// TIA Portal V20 export
// export: Created 2026-10-20T12:51:09.2669842Z, ExportSetting WithDefaults, DisplayName Totally Integrated Automation Portal, DisplayVersion V20 Update 6, DisplayName TIA Portal Openness, DisplayVersion V20 Update 6, DisplayName TIA Portal Version Control Interface, DisplayVersion V20 Update 6, DisplayName SINAMICS Startdrive Advanced, DisplayVersion V20 SP1, DisplayName SINAMICS Startdrive G130, G150, S120, S150, SINAMICS MV, G220, S200, S210, DisplayVersion V20 SP1, DisplayName SINAMICS Startdrive G110M, G120, G120C, G120D, G120P, G115D, DisplayVersion V20 SP1, DisplayName STEP 7 Professional, DisplayVersion V20 Update 6, DisplayName STEP 7 Safety, DisplayVersion V20 Update 2, DisplayName WinCC Basic/Comfort/Advanced, DisplayVersion V20 Update 6, DisplayName WinCC Unified, DisplayVersion V20 Update 6
FUNCTION_BLOCK "Remote_Panel"   // FB17, F_LAD
{ S7_Optimized_Access := 'TRUE' }
VERSION : 0.1
// stored: AutoNumber true, IsIECCheckEnabled false, UDAEnableTagReadback false
   VAR_INPUT
      ID : Int;
      Overtravel_Lower_limit : Bool;
      Overtravel_Upper_limit : Bool;
      Estop : Bool;
      Reset : Bool;
      Chain_Slack_1 : Bool;
      Chain_Slack_2 : Bool;
      Chain_Slack_3 : Bool;
      Chain_Slack_4 : Bool;
      "Light Guards CX101" : Bool;
      "Light Guards CX201" : Bool;
      Gate_1 : Bool;
      Gate_2 : Bool;
      EStop_Lock_1 : Bool;
      EStop_Lock_2 : Bool;
      Lock_Secured_1 : Bool;
      Lock_Secured_2 : Bool;
      "EStop Level 1" : Bool;
      "EStop Level 2" : Bool;
      "EStop Level 3" : Bool;
      "EStop Level 4" : Bool;
      "EStop Level 5" : Bool;
      "EStop Level 6" : Bool;
      "EStop Level 7" : Bool;
      "EStop Level 8" : Bool;
      Bypass : "F_Bypass_RemotePanel";
      Material_Selection_1 : Bool;
      MR_1 : Bool;
      Material_Selection_2 : Bool;
      MR_2 : Bool;
      Overhang_Left : Bool;
      Overhang_Right : Bool;
   END_VAR
   VAR_OUTPUT
      Safety_OK : Bool;
      Bypass_Warning : Bool;
      "STO VTD - CH1" : Bool;
      "STO VTD - CH2" : Bool;
      "STO CONVEYOR VTD - CH1" : Bool;
      "STO CONVEYOR VTD - CH2" : Bool;
      "STO CNV VFD (Level 1,2,3 - Side1) - CH1" : Bool;
      "STO CNV VFD (Level 1,2,3 - Side1) - CH2" : Bool;
      "STO CNV VFD (Level 1,2,3 - Side2) - CH1" : Bool;
      "STO CNV VFD (Level 1,2,3 - Side2) - CH2" : Bool;
      "STO CNV VFD (Level 4,5,6 - Side1) - CH1" : Bool;
      "STO CNV VFD (Level 4,5,6 - Side1) - CH2" : Bool;
      "STO CNV VFD (Level 4,5,6 - Side2) - CH1" : Bool;
      "STO CNV VFD (Level 4,5,6 - Side2) - CH2" : Bool;
      "STO CNV VFD (Level 7,8 - Side1) - CH1" : Bool;
      "STO CNV VFD (Level 7,8 - Side1) - CH2" : Bool;
      "STO CNV VFD (Level 7,8 - Side2) - CH1" : Bool;
      "STO CNV VFD (Level 7,8 - Side2) - CH2" : Bool;
      "Power Enable Safety Stopper Conveyors (Level 1,2,3 - Side1) - CH1" : Bool;
      "Power Enable Safety Stopper Conveyors (Level 1,2,3 - Side1) - CH2" : Bool;
      "Power Enable Safety Stopper Conveyors (Level 1,2,3 - Side2) - CH1" : Bool;
      "Power Enable Safety Stopper Conveyors (Level 1,2,3 - Side2) - CH2" : Bool;
      "Power Enable Safety Stopper Conveyors (Level 4,5,6 - Side1) - CH1" : Bool;
      "Power Enable Safety Stopper Conveyors (Level 4,5,6 - Side1) - CH2" : Bool;
      "Power Enable Safety Stopper Conveyors (Level 4,5,6 - Side2) - CH1" : Bool;
      "Power Enable Safety Stopper Conveyors (Level 4,5,6 - Side2) - CH2" : Bool;
      "Power Enable Safety Stopper Conveyors (Level 7,8 - Side1) - CH1" : Bool;
      "Power Enable Safety Stopper Conveyors (Level 7,8 - Side1) - CH2" : Bool;
      "Power Enable Safety Stopper Conveyors (Level 7,8 - Side2) - CH1" : Bool;
      "Power Enable Safety Stopper Conveyors (Level 7,8 - Side2) - CH2" : Bool;
      "VTU Hoist Brake Sfty Enable - CH1" : Bool;
      "VTU Hoist Brake Sfty Enable - CH2" : Bool;
      ACK { ExternalAccessible := 'False'; ExternalVisible := 'False'; ExternalWritable := 'False'} : Bool;
      L1_OK : Bool;
      L2_OK : Bool;
      L3_OK : Bool;
      L4_OK : Bool;
      L5_OK : Bool;
      L6_OK : Bool;
      L7_OK : Bool;
      L8_OK : Bool;
      EStop_Lock_1_OK : Bool;
      EStop_Lock_2_OK : Bool;
      Lock_Secured_1_OK : Bool;
      Lock_Secured_2_OK : Bool;
      Safety_Ok_Conf : Bool;
   END_VAR
   VAR
      Overtravel_Lower_Limit_DB : ESTOP1;
      Overtravel_Upper_Limit_DB : ESTOP1;
      Estop_Cabinet_DB : ESTOP1;
      Chain_Slack_1_DB : ESTOP1;
      Chain_Slack_2_DB : ESTOP1;
      Chain_Slack_3_DB : ESTOP1;
      Chain_Slack_4_DB : ESTOP1;
      Light_Guards_CX101 : ESTOP1;
      Light_Guards_CX201 : ESTOP1;
      Gate_1_DB : ESTOP1;
      Gate_2_DB : ESTOP1;
      EStop_Lock_1_DB : ESTOP1;
      EStop_Lock_2_DB : ESTOP1;
      Lock_Secured_1_DB : ESTOP1;
      Lock_Secured_2_DB : ESTOP1;
      "EStop Level 1_DB" : ESTOP1;
      "EStop Level 2_DB" : ESTOP1;
      "EStop Level 3_DB" : ESTOP1;
      "EStop Level 4_DB" : ESTOP1;
      "EStop Level 5_DB" : ESTOP1;
      "EStop Level 6_DB" : ESTOP1;
      "EStop Level 7_DB" : ESTOP1;
      "EStop Level 8_DB" : ESTOP1;
      Mute_LG_1_DB : "SICK Safe Entry Exit HW PLC V02";
      Distance_Materia_To_LG : DInt;
      Mute_LG_2_DB : "SICK Safe Entry Exit HW PLC V02";
      F_T_Delay_Sae_OK : TOF;
      F_T_Delay_CL_4 : TOF;
      F_T_Delay_CL_3 : TOF;
      F_T_Delay_CL_2 : TOF;
      F_T_Delay_CL_1 : TOF;
      Chain_Slack_1_Filtered { ExternalAccessible := 'False'; ExternalVisible := 'False'; ExternalWritable := 'False'} : Bool;
      Chain_Slack_2_Filtered { ExternalAccessible := 'False'; ExternalVisible := 'False'; ExternalWritable := 'False'} : Bool;
      Chain_Slack_3_Filtered { ExternalAccessible := 'False'; ExternalVisible := 'False'; ExternalWritable := 'False'} : Bool;
      Chain_Slack_4_Filtered { ExternalAccessible := 'False'; ExternalVisible := 'False'; ExternalWritable := 'False'} : Bool;
      Light_Guard_Tuned : Bool;
      Light_Guard_Tuned_Euro : Bool;
      Light_Guard_Tuned_UK : Bool;
      Light_Guard_Tuned_UK_Infeed : Bool;
      Light_Guard_Tuned_Euro_Infeed : Bool;
      Light_Guard_Tuned_Infeed : Bool;
      F_Timer_Infeed_UK : TP;
      F_Timer_Infeed_E : TP;
      F_Timer_Outfeed_UK : TP;
      F_Timer_Outfeed_E : TP;
      Overhang_Left_DB : ESTOP1;
      Overhang_Right_DB : ESTOP1;
   END_VAR
   VAR_TEMP
      EStop_Levels_OK : Bool;
   END_VAR
   VAR_TEMP   // added for the SCL form of the ladder/FBD networks
      _w1 : Bool;
   END_VAR
BEGIN

REGION Network 1: RESET CABINET
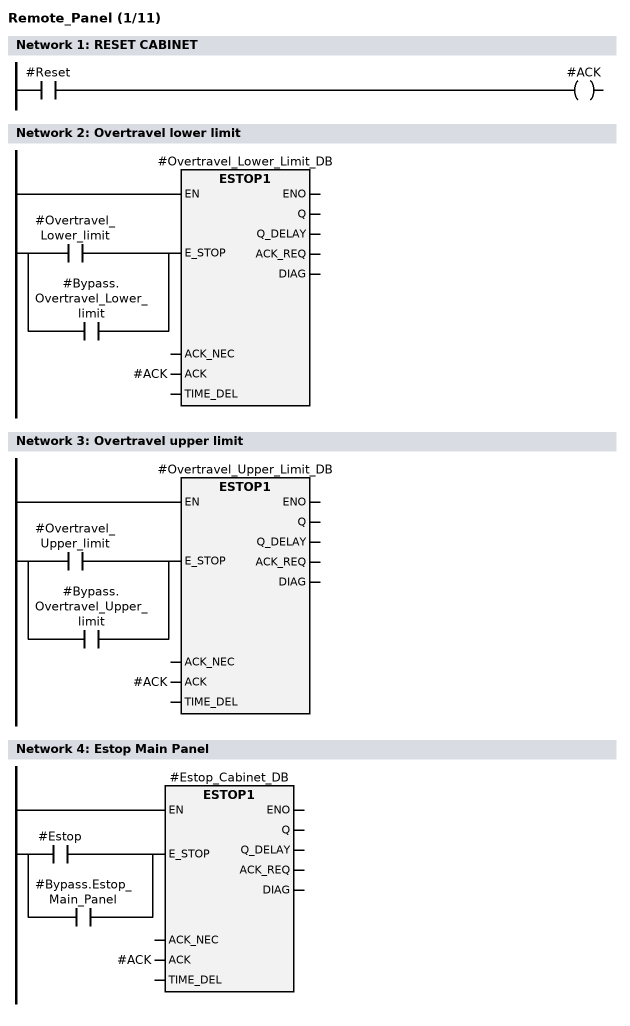
   RUNG wire#powerrail
      Contact( #Reset )
      Coil( #ACK )
   END_RUNG
   // the same network as SCL:
   #ACK := #Reset;
END_REGION

REGION Network 2: Overtravel lower limit
   RUNG wire#powerrail
      #Overtravel_Lower_Limit_DB.ESTOP1(E_STOP := wire#w1, ACK_NEC :=, ACK := #ACK, TIME_DEL :=, Q =>, Q_DELAY =>, ACK_REQ =>, DIAG =>)
   END_RUNG
   RUNG wire#powerrail
      Contact( #Overtravel_Lower_limit )
   END_RUNG wire#w1
   RUNG wire#powerrail
      Contact( #Bypass.Overtravel_Lower_limit )
   END_RUNG wire#w1
   // the same network as SCL:
   #Overtravel_Lower_Limit_DB(E_STOP := #Overtravel_Lower_limit OR #Bypass.Overtravel_Lower_limit, ACK := #ACK);   // ESTOP1
END_REGION

REGION Network 3: Overtravel upper limit
   RUNG wire#powerrail
      #Overtravel_Upper_Limit_DB.ESTOP1(E_STOP := wire#w1, ACK_NEC :=, ACK := #ACK, TIME_DEL :=, Q =>, Q_DELAY =>, ACK_REQ =>, DIAG =>)
   END_RUNG
   RUNG wire#powerrail
      Contact( #Overtravel_Upper_limit )
   END_RUNG wire#w1
   RUNG wire#powerrail
      Contact( #Bypass.Overtravel_Upper_limit )
   END_RUNG wire#w1
   // the same network as SCL:
   #Overtravel_Upper_Limit_DB(E_STOP := #Overtravel_Upper_limit OR #Bypass.Overtravel_Upper_limit, ACK := #ACK);   // ESTOP1
END_REGION

REGION Network 4: Estop Main Panel
   RUNG wire#powerrail
      #Estop_Cabinet_DB.ESTOP1(E_STOP := wire#w1, ACK_NEC :=, ACK := #ACK, TIME_DEL :=, Q =>, Q_DELAY =>, ACK_REQ =>, DIAG =>)
   END_RUNG
   RUNG wire#powerrail
      Contact( #Estop )
   END_RUNG wire#w1
   RUNG wire#powerrail
      Contact( #Bypass.Estop_Main_Panel )
   END_RUNG wire#w1
   // the same network as SCL:
   #Estop_Cabinet_DB(E_STOP := #Estop OR #Bypass.Estop_Main_Panel, ACK := #ACK);   // ESTOP1
END_REGION

REGION Network 5: Chain slack 1
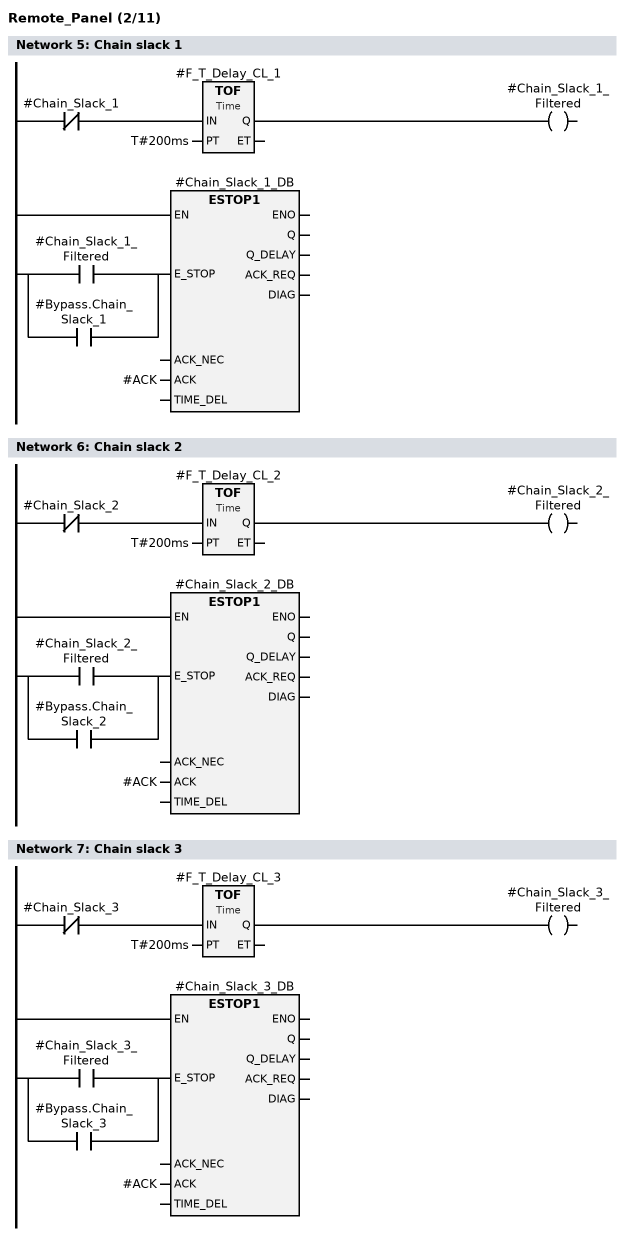
   RUNG wire#powerrail
      I_Contact( #Chain_Slack_1 )
      { S7_Templates := "[time_type := Time, codedbool_type := DInt]" } #F_T_Delay_CL_1.TOF(pt := T#200ms, et =>)
      Coil( #Chain_Slack_1_Filtered )
   END_RUNG
   RUNG wire#powerrail
      #Chain_Slack_1_DB.ESTOP1(E_STOP := wire#w1, ACK_NEC :=, ACK := #ACK, TIME_DEL :=, Q =>, Q_DELAY =>, ACK_REQ =>, DIAG =>)
   END_RUNG
   RUNG wire#powerrail
      Contact( #Chain_Slack_1_Filtered )
   END_RUNG wire#w1
   RUNG wire#powerrail
      Contact( #Bypass.Chain_Slack_1 )
   END_RUNG wire#w1
   // the same network as SCL:
   #F_T_Delay_CL_1.TOF(IN := NOT #Chain_Slack_1, PT := T#200ms);
   #Chain_Slack_1_Filtered := #F_T_Delay_CL_1.Q;
   #Chain_Slack_1_DB(E_STOP := #Chain_Slack_1_Filtered OR #Bypass.Chain_Slack_1, ACK := #ACK);   // ESTOP1
END_REGION

REGION Network 6: Chain slack 2
   RUNG wire#powerrail
      I_Contact( #Chain_Slack_2 )
      { S7_Templates := "[time_type := Time, codedbool_type := DInt]" } #F_T_Delay_CL_2.TOF(pt := T#200ms, et =>)
      Coil( #Chain_Slack_2_Filtered )
   END_RUNG
   RUNG wire#powerrail
      #Chain_Slack_2_DB.ESTOP1(E_STOP := wire#w1, ACK_NEC :=, ACK := #ACK, TIME_DEL :=, Q =>, Q_DELAY =>, ACK_REQ =>, DIAG =>)
   END_RUNG
   RUNG wire#powerrail
      Contact( #Chain_Slack_2_Filtered )
   END_RUNG wire#w1
   RUNG wire#powerrail
      Contact( #Bypass.Chain_Slack_2 )
   END_RUNG wire#w1
   // the same network as SCL:
   #F_T_Delay_CL_2.TOF(IN := NOT #Chain_Slack_2, PT := T#200ms);
   #Chain_Slack_2_Filtered := #F_T_Delay_CL_2.Q;
   #Chain_Slack_2_DB(E_STOP := #Chain_Slack_2_Filtered OR #Bypass.Chain_Slack_2, ACK := #ACK);   // ESTOP1
END_REGION

REGION Network 7: Chain slack 3
   RUNG wire#powerrail
      I_Contact( #Chain_Slack_3 )
      { S7_Templates := "[time_type := Time, codedbool_type := DInt]" } #F_T_Delay_CL_3.TOF(pt := T#200ms, et =>)
      Coil( #Chain_Slack_3_Filtered )
   END_RUNG
   RUNG wire#powerrail
      #Chain_Slack_3_DB.ESTOP1(E_STOP := wire#w1, ACK_NEC :=, ACK := #ACK, TIME_DEL :=, Q =>, Q_DELAY =>, ACK_REQ =>, DIAG =>)
   END_RUNG
   RUNG wire#powerrail
      Contact( #Chain_Slack_3_Filtered )
   END_RUNG wire#w1
   RUNG wire#powerrail
      Contact( #Bypass.Chain_Slack_3 )
   END_RUNG wire#w1
   // the same network as SCL:
   #F_T_Delay_CL_3.TOF(IN := NOT #Chain_Slack_3, PT := T#200ms);
   #Chain_Slack_3_Filtered := #F_T_Delay_CL_3.Q;
   #Chain_Slack_3_DB(E_STOP := #Chain_Slack_3_Filtered OR #Bypass.Chain_Slack_3, ACK := #ACK);   // ESTOP1
END_REGION

REGION Network 8: Chain slack 4
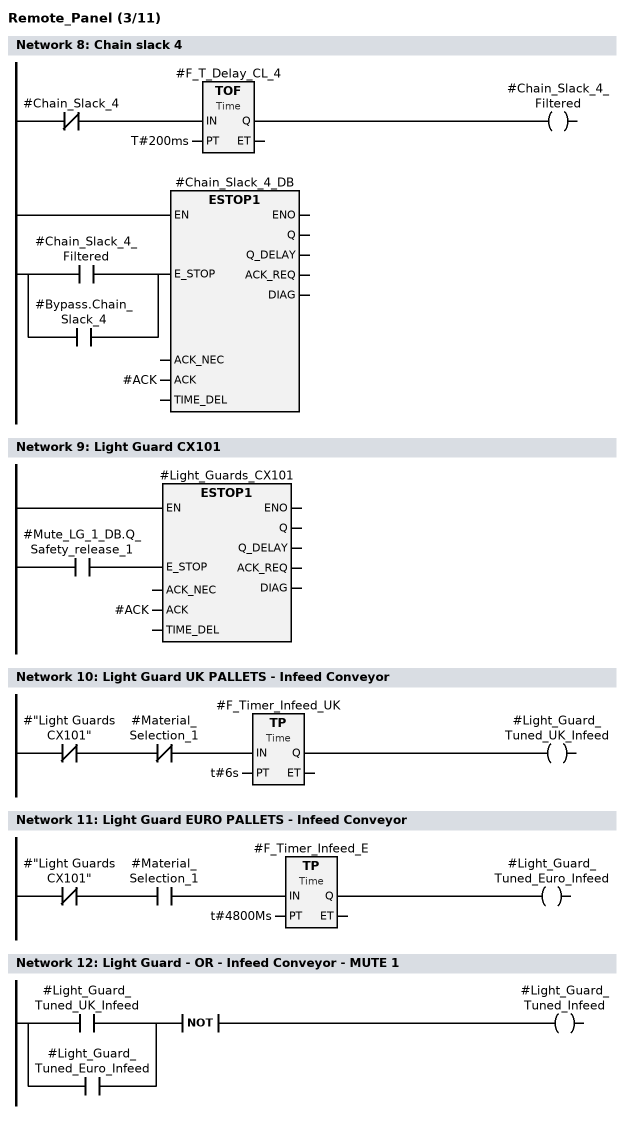
   RUNG wire#powerrail
      I_Contact( #Chain_Slack_4 )
      { S7_Templates := "[time_type := Time, codedbool_type := DInt]" } #F_T_Delay_CL_4.TOF(pt := T#200ms, et =>)
      Coil( #Chain_Slack_4_Filtered )
   END_RUNG
   RUNG wire#powerrail
      #Chain_Slack_4_DB.ESTOP1(E_STOP := wire#w1, ACK_NEC :=, ACK := #ACK, TIME_DEL :=, Q =>, Q_DELAY =>, ACK_REQ =>, DIAG =>)
   END_RUNG
   RUNG wire#powerrail
      Contact( #Chain_Slack_4_Filtered )
   END_RUNG wire#w1
   RUNG wire#powerrail
      Contact( #Bypass.Chain_Slack_4 )
   END_RUNG wire#w1
   // the same network as SCL:
   #F_T_Delay_CL_4.TOF(IN := NOT #Chain_Slack_4, PT := T#200ms);
   #Chain_Slack_4_Filtered := #F_T_Delay_CL_4.Q;
   #Chain_Slack_4_DB(E_STOP := #Chain_Slack_4_Filtered OR #Bypass.Chain_Slack_4, ACK := #ACK);   // ESTOP1
END_REGION

REGION Network 9: Light Guard CX101
   RUNG wire#powerrail
      #Light_Guards_CX101.ESTOP1(E_STOP := wire#w1, ACK_NEC :=, ACK := #ACK, TIME_DEL :=, Q =>, Q_DELAY =>, ACK_REQ =>, DIAG =>)
   END_RUNG
   RUNG wire#powerrail
      Contact( #Mute_LG_1_DB.Q_Safety_release_1 )
   END_RUNG wire#w1
   // the same network as SCL:
   #Light_Guards_CX101(E_STOP := #Mute_LG_1_DB.Q_Safety_release_1, ACK := #ACK);   // ESTOP1
END_REGION

REGION Network 10: Light Guard UK PALLETS - Infeed Conveyor
   RUNG wire#powerrail
      I_Contact( #"Light Guards CX101" )
      I_Contact( #Material_Selection_1 )
      { S7_Templates := "[time_type := Time, codedbool_type := DInt]" } #F_Timer_Infeed_UK.TP(pt := t#6s, et =>)
      Coil( #Light_Guard_Tuned_UK_Infeed )
   END_RUNG
   // the same network as SCL:
   #F_Timer_Infeed_UK.TP(IN := NOT #"Light Guards CX101" AND NOT #Material_Selection_1, PT := t#6s);
   #Light_Guard_Tuned_UK_Infeed := #F_Timer_Infeed_UK.Q;
END_REGION

REGION Network 11: Light Guard EURO PALLETS - Infeed Conveyor
   RUNG wire#powerrail
      I_Contact( #"Light Guards CX101" )
      Contact( #Material_Selection_1 )
      { S7_Templates := "[time_type := Time, codedbool_type := DInt]" } #F_Timer_Infeed_E.TP(pt := t#4800Ms, et =>)
      Coil( #Light_Guard_Tuned_Euro_Infeed )
   END_RUNG
   // the same network as SCL:
   #F_Timer_Infeed_E.TP(IN := NOT #"Light Guards CX101" AND #Material_Selection_1, PT := t#4800Ms);
   #Light_Guard_Tuned_Euro_Infeed := #F_Timer_Infeed_E.Q;
END_REGION

REGION Network 12: Light Guard - OR - Infeed Conveyor - MUTE 1
   RUNG wire#powerrail
      Contact( #Light_Guard_Tuned_UK_Infeed )
      wire#w1
      Not()
      Coil( #Light_Guard_Tuned_Infeed )
   END_RUNG
   RUNG wire#powerrail
      Contact( #Light_Guard_Tuned_Euro_Infeed )
   END_RUNG wire#w1
   // the same network as SCL:
   #Light_Guard_Tuned_Infeed := NOT (#Light_Guard_Tuned_UK_Infeed OR #Light_Guard_Tuned_Euro_Infeed);
END_REGION

REGION Network 13: MUTE 1
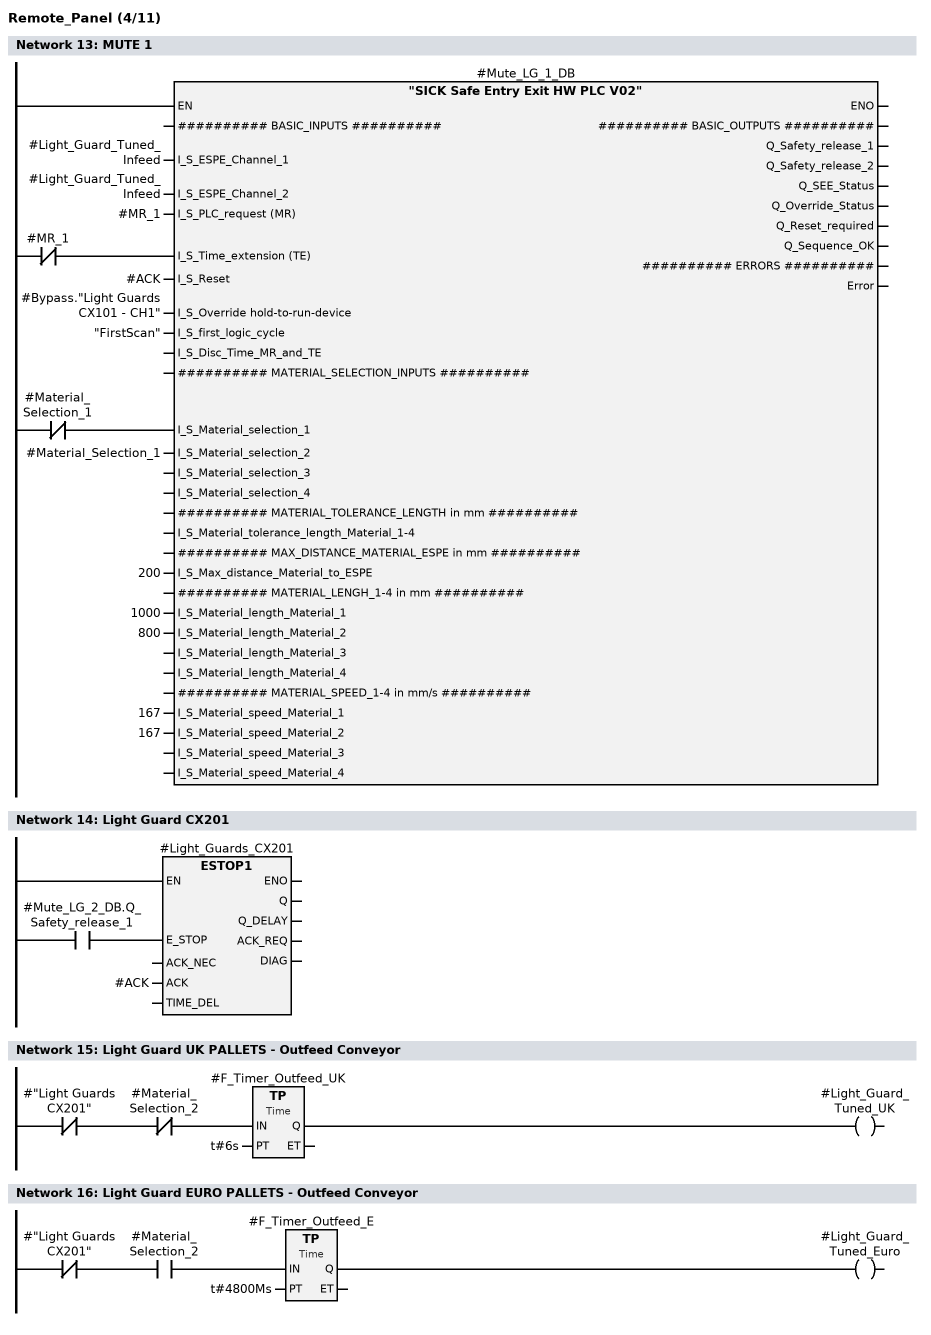
   RUNG wire#powerrail
      #Mute_LG_1_DB("I_S_Time_extension (TE)" := wire#w1, I_S_Material_selection_1 := wire#w2, "########## BASIC_INPUTS ##########" :=, I_S_ESPE_Channel_1 := #Light_Guard_Tuned_Infeed, I_S_ESPE_Channel_2 := #Light_Guard_Tuned_Infeed, "I_S_PLC_request (MR)" := #MR_1, I_S_Reset := #ACK, "I_S_Override hold-to-run-device" := #Bypass."Light Guards CX101 - CH1", I_S_first_logic_cycle := "FirstScan", I_S_Disc_Time_MR_and_TE :=, "########## MATERIAL_SELECTION_INPUTS ##########" :=, I_S_Material_selection_2 := #Material_Selection_1, I_S_Material_selection_3 :=, I_S_Material_selection_4 :=, "########## MATERIAL_TOLERANCE_LENGTH in mm ##########" :=, "I_S_Material_tolerance_length_Material_1-4" :=, "########## MAX_DISTANCE_MATERIAL_ESPE in mm ##########" :=, I_S_Max_distance_Material_to_ESPE := 200, "########## MATERIAL_LENGH_1-4 in mm ##########" :=, I_S_Material_length_Material_1 := 1000, I_S_Material_length_Material_2 := 800, I_S_Material_length_Material_3 :=, I_S_Material_length_Material_4 :=, "########## MATERIAL_SPEED_1-4 in mm/s ##########" :=, I_S_Material_speed_Material_1 := 167, I_S_Material_speed_Material_2 := 167, I_S_Material_speed_Material_3 :=, I_S_Material_speed_Material_4 :=, "########## BASIC_OUTPUTS ##########" =>, Q_Safety_release_1 =>, Q_Safety_release_2 =>, Q_SEE_Status =>, Q_Override_Status =>, Q_Reset_required =>, Q_Sequence_OK =>, "########## ERRORS ##########" =>, Error =>)
   END_RUNG
   RUNG wire#powerrail
      I_Contact( #MR_1 )
   END_RUNG wire#w1
   RUNG wire#powerrail
      I_Contact( #Material_Selection_1 )
   END_RUNG wire#w2
   // the same network as SCL:
   #Mute_LG_1_DB(I_S_ESPE_Channel_1 := #Light_Guard_Tuned_Infeed,   // "SICK Safe Entry Exit HW PLC V02"
                 I_S_ESPE_Channel_2 := #Light_Guard_Tuned_Infeed,
                 "I_S_PLC_request (MR)" := #MR_1,
                 "I_S_Time_extension (TE)" := NOT #MR_1,
                 I_S_Reset := #ACK,
                 "I_S_Override hold-to-run-device" := #Bypass."Light Guards CX101 - CH1",
                 I_S_first_logic_cycle := "FirstScan",
                 I_S_Material_selection_1 := NOT #Material_Selection_1,
                 I_S_Material_selection_2 := #Material_Selection_1,
                 I_S_Max_distance_Material_to_ESPE := 200,
                 I_S_Material_length_Material_1 := 1000,
                 I_S_Material_length_Material_2 := 800,
                 I_S_Material_speed_Material_1 := 167,
                 I_S_Material_speed_Material_2 := 167);
END_REGION

REGION Network 14: Light Guard CX201
   RUNG wire#powerrail
      #Light_Guards_CX201.ESTOP1(E_STOP := wire#w1, ACK_NEC :=, ACK := #ACK, TIME_DEL :=, Q =>, Q_DELAY =>, ACK_REQ =>, DIAG =>)
   END_RUNG
   RUNG wire#powerrail
      Contact( #Mute_LG_2_DB.Q_Safety_release_1 )
   END_RUNG wire#w1
   // the same network as SCL:
   #Light_Guards_CX201(E_STOP := #Mute_LG_2_DB.Q_Safety_release_1, ACK := #ACK);   // ESTOP1
END_REGION

REGION Network 15: Light Guard UK PALLETS - Outfeed Conveyor
   RUNG wire#powerrail
      I_Contact( #"Light Guards CX201" )
      I_Contact( #Material_Selection_2 )
      { S7_Templates := "[time_type := Time, codedbool_type := DInt]" } #F_Timer_Outfeed_UK.TP(pt := t#6s, et =>)
      Coil( #Light_Guard_Tuned_UK )
   END_RUNG
   // the same network as SCL:
   #F_Timer_Outfeed_UK.TP(IN := NOT #"Light Guards CX201" AND NOT #Material_Selection_2, PT := t#6s);
   #Light_Guard_Tuned_UK := #F_Timer_Outfeed_UK.Q;
END_REGION

REGION Network 16: Light Guard EURO PALLETS - Outfeed Conveyor
   RUNG wire#powerrail
      I_Contact( #"Light Guards CX201" )
      Contact( #Material_Selection_2 )
      { S7_Templates := "[time_type := Time, codedbool_type := DInt]" } #F_Timer_Outfeed_E.TP(pt := t#4800Ms, et =>)
      Coil( #Light_Guard_Tuned_Euro )
   END_RUNG
   // the same network as SCL:
   #F_Timer_Outfeed_E.TP(IN := NOT #"Light Guards CX201" AND #Material_Selection_2, PT := t#4800Ms);
   #Light_Guard_Tuned_Euro := #F_Timer_Outfeed_E.Q;
END_REGION

REGION Network 17: Light Guard - OR - Infeed Conveyor - MUTE 2
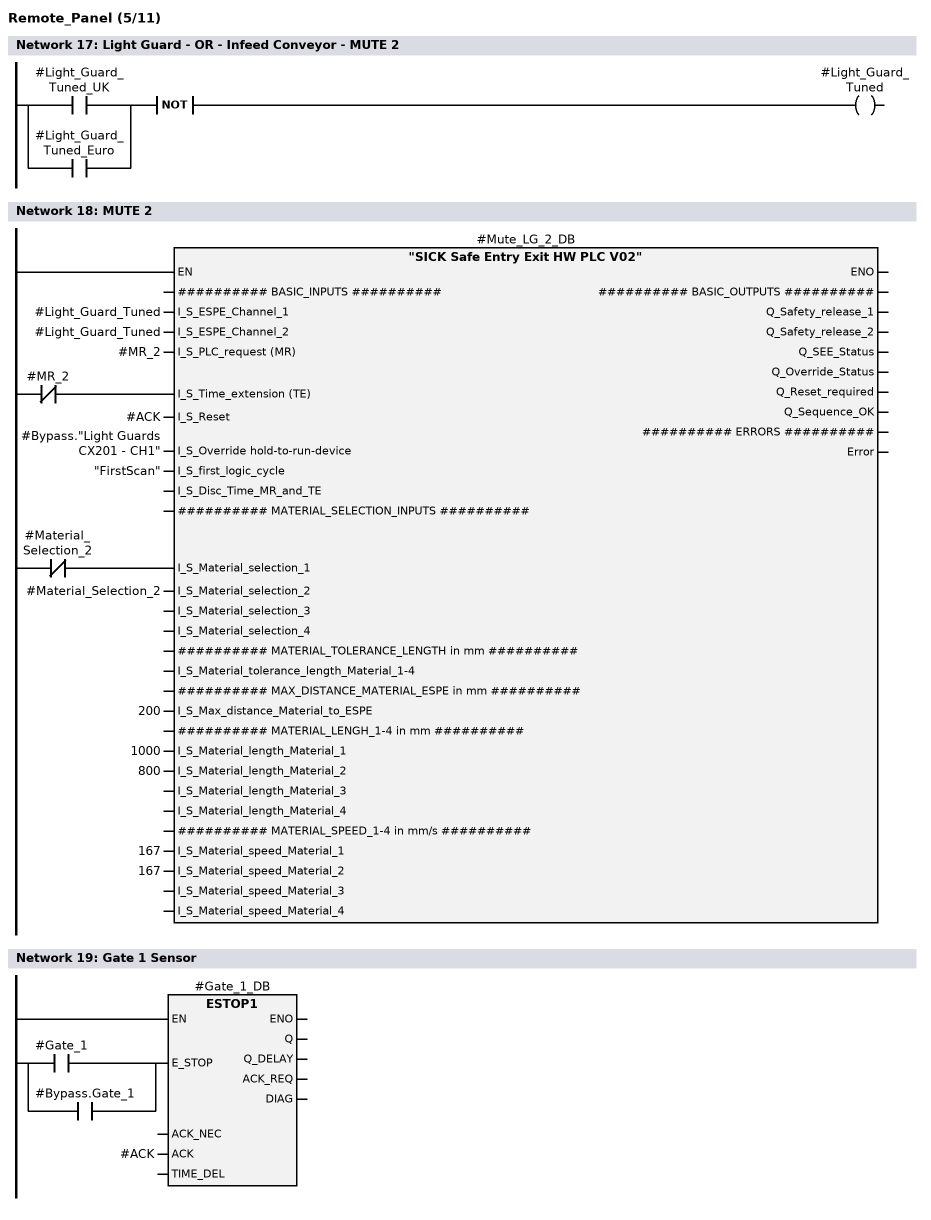
   RUNG wire#powerrail
      Contact( #Light_Guard_Tuned_UK )
      wire#w1
      Not()
      Coil( #Light_Guard_Tuned )
   END_RUNG
   RUNG wire#powerrail
      Contact( #Light_Guard_Tuned_Euro )
   END_RUNG wire#w1
   // the same network as SCL:
   #Light_Guard_Tuned := NOT (#Light_Guard_Tuned_UK OR #Light_Guard_Tuned_Euro);
END_REGION

REGION Network 18: MUTE 2
   RUNG wire#powerrail
      #Mute_LG_2_DB("I_S_Time_extension (TE)" := wire#w1, I_S_Material_selection_1 := wire#w2, "########## BASIC_INPUTS ##########" :=, I_S_ESPE_Channel_1 := #Light_Guard_Tuned, I_S_ESPE_Channel_2 := #Light_Guard_Tuned, "I_S_PLC_request (MR)" := #MR_2, I_S_Reset := #ACK, "I_S_Override hold-to-run-device" := #Bypass."Light Guards CX201 - CH1", I_S_first_logic_cycle := "FirstScan", I_S_Disc_Time_MR_and_TE :=, "########## MATERIAL_SELECTION_INPUTS ##########" :=, I_S_Material_selection_2 := #Material_Selection_2, I_S_Material_selection_3 :=, I_S_Material_selection_4 :=, "########## MATERIAL_TOLERANCE_LENGTH in mm ##########" :=, "I_S_Material_tolerance_length_Material_1-4" :=, "########## MAX_DISTANCE_MATERIAL_ESPE in mm ##########" :=, I_S_Max_distance_Material_to_ESPE := 200, "########## MATERIAL_LENGH_1-4 in mm ##########" :=, I_S_Material_length_Material_1 := 1000, I_S_Material_length_Material_2 := 800, I_S_Material_length_Material_3 :=, I_S_Material_length_Material_4 :=, "########## MATERIAL_SPEED_1-4 in mm/s ##########" :=, I_S_Material_speed_Material_1 := 167, I_S_Material_speed_Material_2 := 167, I_S_Material_speed_Material_3 :=, I_S_Material_speed_Material_4 :=, "########## BASIC_OUTPUTS ##########" =>, Q_Safety_release_1 =>, Q_Safety_release_2 =>, Q_SEE_Status =>, Q_Override_Status =>, Q_Reset_required =>, Q_Sequence_OK =>, "########## ERRORS ##########" =>, Error =>)
   END_RUNG
   RUNG wire#powerrail
      I_Contact( #MR_2 )
   END_RUNG wire#w1
   RUNG wire#powerrail
      I_Contact( #Material_Selection_2 )
   END_RUNG wire#w2
   // the same network as SCL:
   #Mute_LG_2_DB(I_S_ESPE_Channel_1 := #Light_Guard_Tuned,   // "SICK Safe Entry Exit HW PLC V02"
                 I_S_ESPE_Channel_2 := #Light_Guard_Tuned,
                 "I_S_PLC_request (MR)" := #MR_2,
                 "I_S_Time_extension (TE)" := NOT #MR_2,
                 I_S_Reset := #ACK,
                 "I_S_Override hold-to-run-device" := #Bypass."Light Guards CX201 - CH1",
                 I_S_first_logic_cycle := "FirstScan",
                 I_S_Material_selection_1 := NOT #Material_Selection_2,
                 I_S_Material_selection_2 := #Material_Selection_2,
                 I_S_Max_distance_Material_to_ESPE := 200,
                 I_S_Material_length_Material_1 := 1000,
                 I_S_Material_length_Material_2 := 800,
                 I_S_Material_speed_Material_1 := 167,
                 I_S_Material_speed_Material_2 := 167);
END_REGION

REGION Network 19: Gate 1 Sensor
   RUNG wire#powerrail
      #Gate_1_DB.ESTOP1(E_STOP := wire#w1, ACK_NEC :=, ACK := #ACK, TIME_DEL :=, Q =>, Q_DELAY =>, ACK_REQ =>, DIAG =>)
   END_RUNG
   RUNG wire#powerrail
      Contact( #Gate_1 )
   END_RUNG wire#w1
   RUNG wire#powerrail
      Contact( #Bypass.Gate_1 )
   END_RUNG wire#w1
   // the same network as SCL:
   #Gate_1_DB(E_STOP := #Gate_1 OR #Bypass.Gate_1, ACK := #ACK);   // ESTOP1
END_REGION

REGION Network 20: Gate 2 Sensor
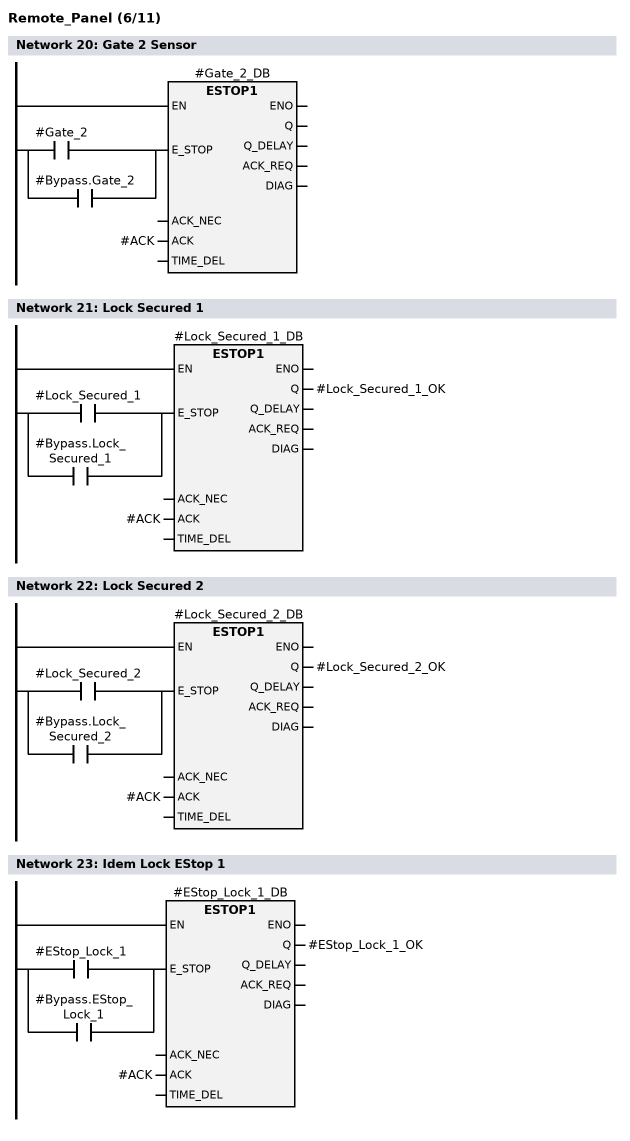
   RUNG wire#powerrail
      #Gate_2_DB.ESTOP1(E_STOP := wire#w1, ACK_NEC :=, ACK := #ACK, TIME_DEL :=, Q =>, Q_DELAY =>, ACK_REQ =>, DIAG =>)
   END_RUNG
   RUNG wire#powerrail
      Contact( #Gate_2 )
   END_RUNG wire#w1
   RUNG wire#powerrail
      Contact( #Bypass.Gate_2 )
   END_RUNG wire#w1
   // the same network as SCL:
   #Gate_2_DB(E_STOP := #Gate_2 OR #Bypass.Gate_2, ACK := #ACK);   // ESTOP1
END_REGION

REGION Network 21: Lock Secured 1
   RUNG wire#powerrail
      #Lock_Secured_1_DB.ESTOP1(E_STOP := wire#w1, ACK_NEC :=, ACK := #ACK, TIME_DEL :=, Q => #Lock_Secured_1_OK, Q_DELAY =>, ACK_REQ =>, DIAG =>)
   END_RUNG
   RUNG wire#powerrail
      Contact( #Lock_Secured_1 )
   END_RUNG wire#w1
   RUNG wire#powerrail
      Contact( #Bypass.Lock_Secured_1 )
   END_RUNG wire#w1
   // the same network as SCL:
   #Lock_Secured_1_DB(E_STOP := #Lock_Secured_1 OR #Bypass.Lock_Secured_1, ACK := #ACK, Q => #Lock_Secured_1_OK);   // ESTOP1
END_REGION

REGION Network 22: Lock Secured 2
   RUNG wire#powerrail
      #Lock_Secured_2_DB.ESTOP1(E_STOP := wire#w1, ACK_NEC :=, ACK := #ACK, TIME_DEL :=, Q => #Lock_Secured_2_OK, Q_DELAY =>, ACK_REQ =>, DIAG =>)
   END_RUNG
   RUNG wire#powerrail
      Contact( #Lock_Secured_2 )
   END_RUNG wire#w1
   RUNG wire#powerrail
      Contact( #Bypass.Lock_Secured_2 )
   END_RUNG wire#w1
   // the same network as SCL:
   #Lock_Secured_2_DB(E_STOP := #Lock_Secured_2 OR #Bypass.Lock_Secured_2, ACK := #ACK, Q => #Lock_Secured_2_OK);   // ESTOP1
END_REGION

REGION Network 23: Idem Lock EStop 1
   RUNG wire#powerrail
      #EStop_Lock_1_DB.ESTOP1(E_STOP := wire#w1, ACK_NEC :=, ACK := #ACK, TIME_DEL :=, Q => #EStop_Lock_1_OK, Q_DELAY =>, ACK_REQ =>, DIAG =>)
   END_RUNG
   RUNG wire#powerrail
      Contact( #EStop_Lock_1 )
   END_RUNG wire#w1
   RUNG wire#powerrail
      Contact( #Bypass.EStop_Lock_1 )
   END_RUNG wire#w1
   // the same network as SCL:
   #EStop_Lock_1_DB(E_STOP := #EStop_Lock_1 OR #Bypass.EStop_Lock_1, ACK := #ACK, Q => #EStop_Lock_1_OK);   // ESTOP1
END_REGION

REGION Network 24: Idem Lock EStop 2
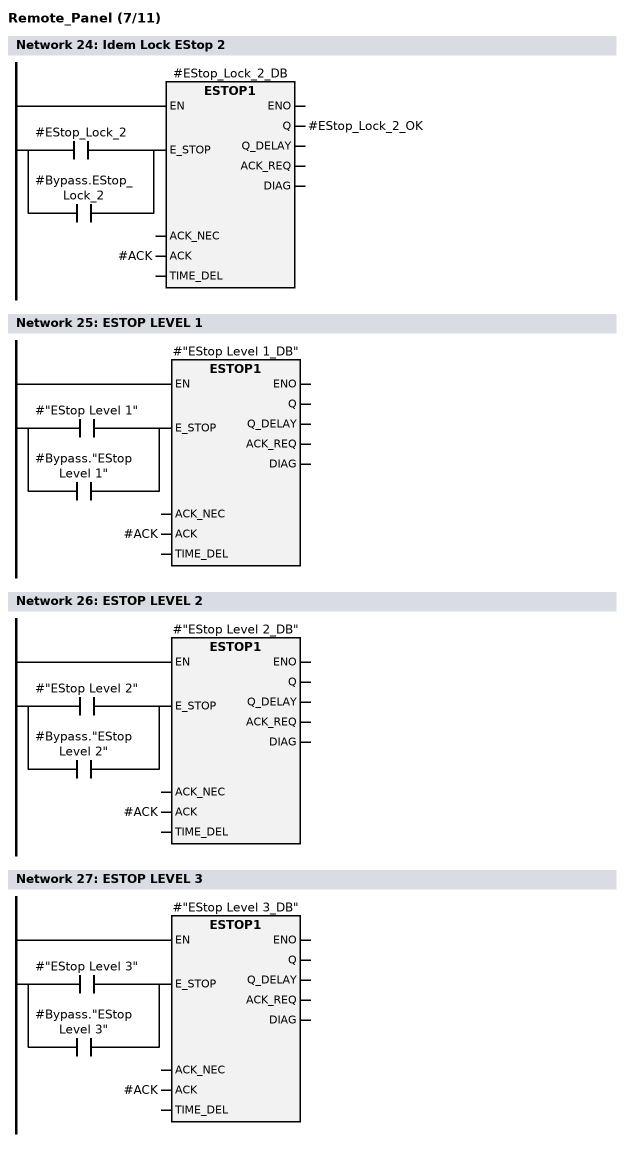
   RUNG wire#powerrail
      #EStop_Lock_2_DB.ESTOP1(E_STOP := wire#w1, ACK_NEC :=, ACK := #ACK, TIME_DEL :=, Q => #EStop_Lock_2_OK, Q_DELAY =>, ACK_REQ =>, DIAG =>)
   END_RUNG
   RUNG wire#powerrail
      Contact( #EStop_Lock_2 )
   END_RUNG wire#w1
   RUNG wire#powerrail
      Contact( #Bypass.EStop_Lock_2 )
   END_RUNG wire#w1
   // the same network as SCL:
   #EStop_Lock_2_DB(E_STOP := #EStop_Lock_2 OR #Bypass.EStop_Lock_2, ACK := #ACK, Q => #EStop_Lock_2_OK);   // ESTOP1
END_REGION

REGION Network 25: ESTOP LEVEL 1
   RUNG wire#powerrail
      #"EStop Level 1_DB".ESTOP1(E_STOP := wire#w1, ACK_NEC :=, ACK := #ACK, TIME_DEL :=, Q =>, Q_DELAY =>, ACK_REQ =>, DIAG =>)
   END_RUNG
   RUNG wire#powerrail
      Contact( #"EStop Level 1" )
   END_RUNG wire#w1
   RUNG wire#powerrail
      Contact( #Bypass."EStop Level 1" )
   END_RUNG wire#w1
   // the same network as SCL:
   #"EStop Level 1_DB"(E_STOP := #"EStop Level 1" OR #Bypass."EStop Level 1", ACK := #ACK);   // ESTOP1
END_REGION

REGION Network 26: ESTOP LEVEL 2
   RUNG wire#powerrail
      #"EStop Level 2_DB".ESTOP1(E_STOP := wire#w1, ACK_NEC :=, ACK := #ACK, TIME_DEL :=, Q =>, Q_DELAY =>, ACK_REQ =>, DIAG =>)
   END_RUNG
   RUNG wire#powerrail
      Contact( #"EStop Level 2" )
   END_RUNG wire#w1
   RUNG wire#powerrail
      Contact( #Bypass."EStop Level 2" )
   END_RUNG wire#w1
   // the same network as SCL:
   #"EStop Level 2_DB"(E_STOP := #"EStop Level 2" OR #Bypass."EStop Level 2", ACK := #ACK);   // ESTOP1
END_REGION

REGION Network 27: ESTOP LEVEL 3
   RUNG wire#powerrail
      #"EStop Level 3_DB".ESTOP1(E_STOP := wire#w1, ACK_NEC :=, ACK := #ACK, TIME_DEL :=, Q =>, Q_DELAY =>, ACK_REQ =>, DIAG =>)
   END_RUNG
   RUNG wire#powerrail
      Contact( #"EStop Level 3" )
   END_RUNG wire#w1
   RUNG wire#powerrail
      Contact( #Bypass."EStop Level 3" )
   END_RUNG wire#w1
   // the same network as SCL:
   #"EStop Level 3_DB"(E_STOP := #"EStop Level 3" OR #Bypass."EStop Level 3", ACK := #ACK);   // ESTOP1
END_REGION

REGION Network 28: ESTOP LEVEL 4
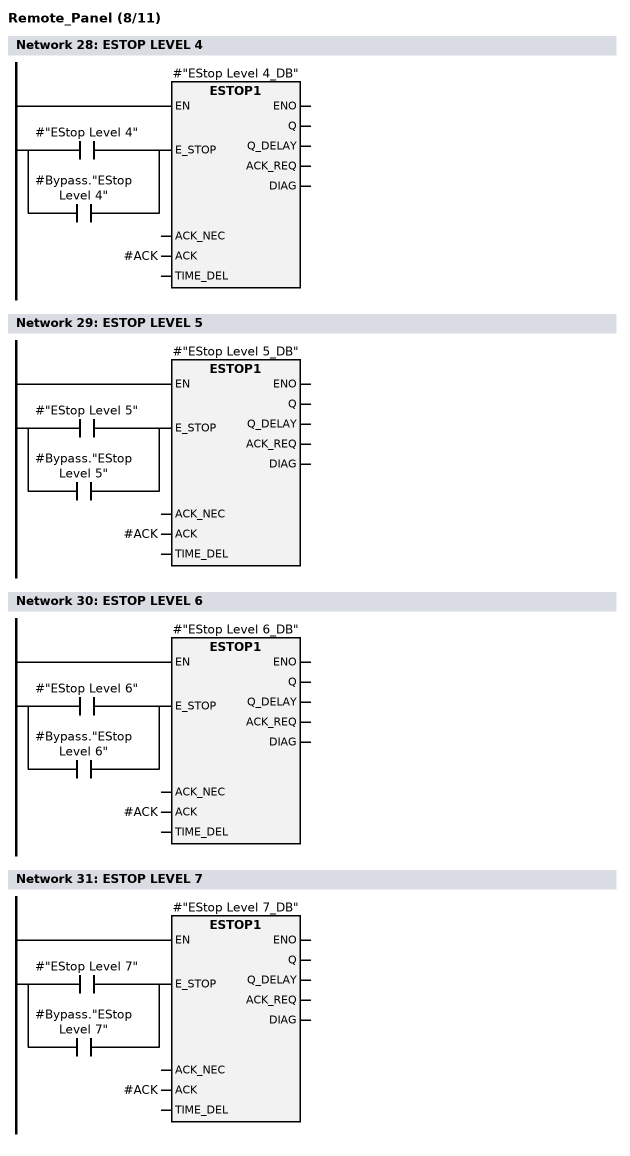
   RUNG wire#powerrail
      #"EStop Level 4_DB".ESTOP1(E_STOP := wire#w1, ACK_NEC :=, ACK := #ACK, TIME_DEL :=, Q =>, Q_DELAY =>, ACK_REQ =>, DIAG =>)
   END_RUNG
   RUNG wire#powerrail
      Contact( #"EStop Level 4" )
   END_RUNG wire#w1
   RUNG wire#powerrail
      Contact( #Bypass."EStop Level 4" )
   END_RUNG wire#w1
   // the same network as SCL:
   #"EStop Level 4_DB"(E_STOP := #"EStop Level 4" OR #Bypass."EStop Level 4", ACK := #ACK);   // ESTOP1
END_REGION

REGION Network 29: ESTOP LEVEL 5
   RUNG wire#powerrail
      #"EStop Level 5_DB".ESTOP1(E_STOP := wire#w1, ACK_NEC :=, ACK := #ACK, TIME_DEL :=, Q =>, Q_DELAY =>, ACK_REQ =>, DIAG =>)
   END_RUNG
   RUNG wire#powerrail
      Contact( #"EStop Level 5" )
   END_RUNG wire#w1
   RUNG wire#powerrail
      Contact( #Bypass."EStop Level 5" )
   END_RUNG wire#w1
   // the same network as SCL:
   #"EStop Level 5_DB"(E_STOP := #"EStop Level 5" OR #Bypass."EStop Level 5", ACK := #ACK);   // ESTOP1
END_REGION

REGION Network 30: ESTOP LEVEL 6
   RUNG wire#powerrail
      #"EStop Level 6_DB".ESTOP1(E_STOP := wire#w1, ACK_NEC :=, ACK := #ACK, TIME_DEL :=, Q =>, Q_DELAY =>, ACK_REQ =>, DIAG =>)
   END_RUNG
   RUNG wire#powerrail
      Contact( #"EStop Level 6" )
   END_RUNG wire#w1
   RUNG wire#powerrail
      Contact( #Bypass."EStop Level 6" )
   END_RUNG wire#w1
   // the same network as SCL:
   #"EStop Level 6_DB"(E_STOP := #"EStop Level 6" OR #Bypass."EStop Level 6", ACK := #ACK);   // ESTOP1
END_REGION

REGION Network 31: ESTOP LEVEL 7
   RUNG wire#powerrail
      #"EStop Level 7_DB".ESTOP1(E_STOP := wire#w1, ACK_NEC :=, ACK := #ACK, TIME_DEL :=, Q =>, Q_DELAY =>, ACK_REQ =>, DIAG =>)
   END_RUNG
   RUNG wire#powerrail
      Contact( #"EStop Level 7" )
   END_RUNG wire#w1
   RUNG wire#powerrail
      Contact( #Bypass."EStop Level 7" )
   END_RUNG wire#w1
   // the same network as SCL:
   #"EStop Level 7_DB"(E_STOP := #"EStop Level 7" OR #Bypass."EStop Level 7", ACK := #ACK);   // ESTOP1
END_REGION

REGION Network 32: ESTOP LEVEL 8
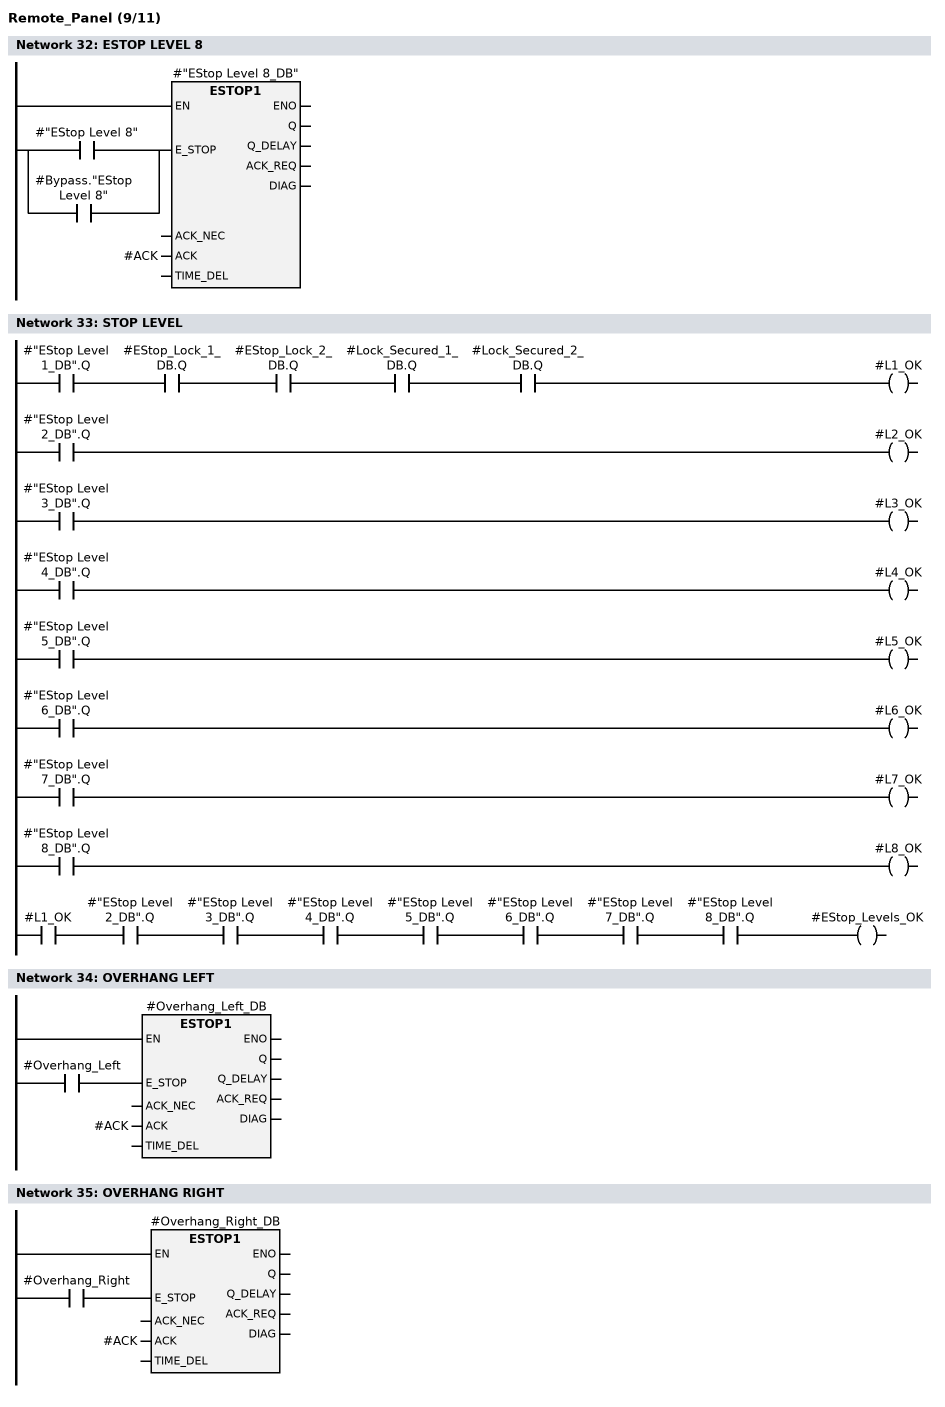
   RUNG wire#powerrail
      #"EStop Level 8_DB".ESTOP1(E_STOP := wire#w1, ACK_NEC :=, ACK := #ACK, TIME_DEL :=, Q =>, Q_DELAY =>, ACK_REQ =>, DIAG =>)
   END_RUNG
   RUNG wire#powerrail
      Contact( #"EStop Level 8" )
   END_RUNG wire#w1
   RUNG wire#powerrail
      Contact( #Bypass."EStop Level 8" )
   END_RUNG wire#w1
   // the same network as SCL:
   #"EStop Level 8_DB"(E_STOP := #"EStop Level 8" OR #Bypass."EStop Level 8", ACK := #ACK);   // ESTOP1
END_REGION

REGION Network 33: STOP LEVEL
   RUNG wire#powerrail
      Contact( #"EStop Level 1_DB".Q )
      Contact( #EStop_Lock_1_DB.Q )
      Contact( #EStop_Lock_2_DB.Q )
      Contact( #Lock_Secured_1_DB.Q )
      Contact( #Lock_Secured_2_DB.Q )
      Coil( #L1_OK )
   END_RUNG
   RUNG wire#powerrail
      Contact( #"EStop Level 2_DB".Q )
      Coil( #L2_OK )
   END_RUNG
   RUNG wire#powerrail
      Contact( #"EStop Level 3_DB".Q )
      Coil( #L3_OK )
   END_RUNG
   RUNG wire#powerrail
      Contact( #"EStop Level 4_DB".Q )
      Coil( #L4_OK )
   END_RUNG
   RUNG wire#powerrail
      Contact( #"EStop Level 5_DB".Q )
      Coil( #L5_OK )
   END_RUNG
   RUNG wire#powerrail
      Contact( #"EStop Level 6_DB".Q )
      Coil( #L6_OK )
   END_RUNG
   RUNG wire#powerrail
      Contact( #"EStop Level 7_DB".Q )
      Coil( #L7_OK )
   END_RUNG
   RUNG wire#powerrail
      Contact( #"EStop Level 8_DB".Q )
      Coil( #L8_OK )
   END_RUNG
   RUNG wire#powerrail
      Contact( #L1_OK )
      Contact( #"EStop Level 2_DB".Q )
      Contact( #"EStop Level 3_DB".Q )
      Contact( #"EStop Level 4_DB".Q )
      Contact( #"EStop Level 5_DB".Q )
      Contact( #"EStop Level 6_DB".Q )
      Contact( #"EStop Level 7_DB".Q )
      Contact( #"EStop Level 8_DB".Q )
      Coil( #EStop_Levels_OK )
   END_RUNG
   // the same network as SCL:
   #L1_OK := #"EStop Level 1_DB".Q AND #EStop_Lock_1_DB.Q AND #EStop_Lock_2_DB.Q AND #Lock_Secured_1_DB.Q AND #Lock_Secured_2_DB.Q;
   #L2_OK := #"EStop Level 2_DB".Q;
   #L3_OK := #"EStop Level 3_DB".Q;
   #L4_OK := #"EStop Level 4_DB".Q;
   #L5_OK := #"EStop Level 5_DB".Q;
   #L6_OK := #"EStop Level 6_DB".Q;
   #L7_OK := #"EStop Level 7_DB".Q;
   #L8_OK := #"EStop Level 8_DB".Q;
   #EStop_Levels_OK := #L1_OK AND #"EStop Level 2_DB".Q AND #"EStop Level 3_DB".Q AND #"EStop Level 4_DB".Q AND #"EStop Level 5_DB".Q AND #"EStop Level 6_DB".Q AND #"EStop Level 7_DB".Q AND #"EStop Level 8_DB".Q;
END_REGION

REGION Network 34: OVERHANG LEFT
   RUNG wire#powerrail
      #Overhang_Left_DB.ESTOP1(E_STOP := wire#w1, ACK_NEC :=, ACK := #ACK, TIME_DEL :=, Q =>, Q_DELAY =>, ACK_REQ =>, DIAG =>)
   END_RUNG
   RUNG wire#powerrail
      Contact( #Overhang_Left )
   END_RUNG wire#w1
   // the same network as SCL:
   #Overhang_Left_DB(E_STOP := #Overhang_Left, ACK := #ACK);   // ESTOP1
END_REGION

REGION Network 35: OVERHANG RIGHT
   RUNG wire#powerrail
      #Overhang_Right_DB.ESTOP1(E_STOP := wire#w1, ACK_NEC :=, ACK := #ACK, TIME_DEL :=, Q =>, Q_DELAY =>, ACK_REQ =>, DIAG =>)
   END_RUNG
   RUNG wire#powerrail
      Contact( #Overhang_Right )
   END_RUNG wire#w1
   // the same network as SCL:
   #Overhang_Right_DB(E_STOP := #Overhang_Right, ACK := #ACK);   // ESTOP1
END_REGION

REGION Network 36: Safety OK
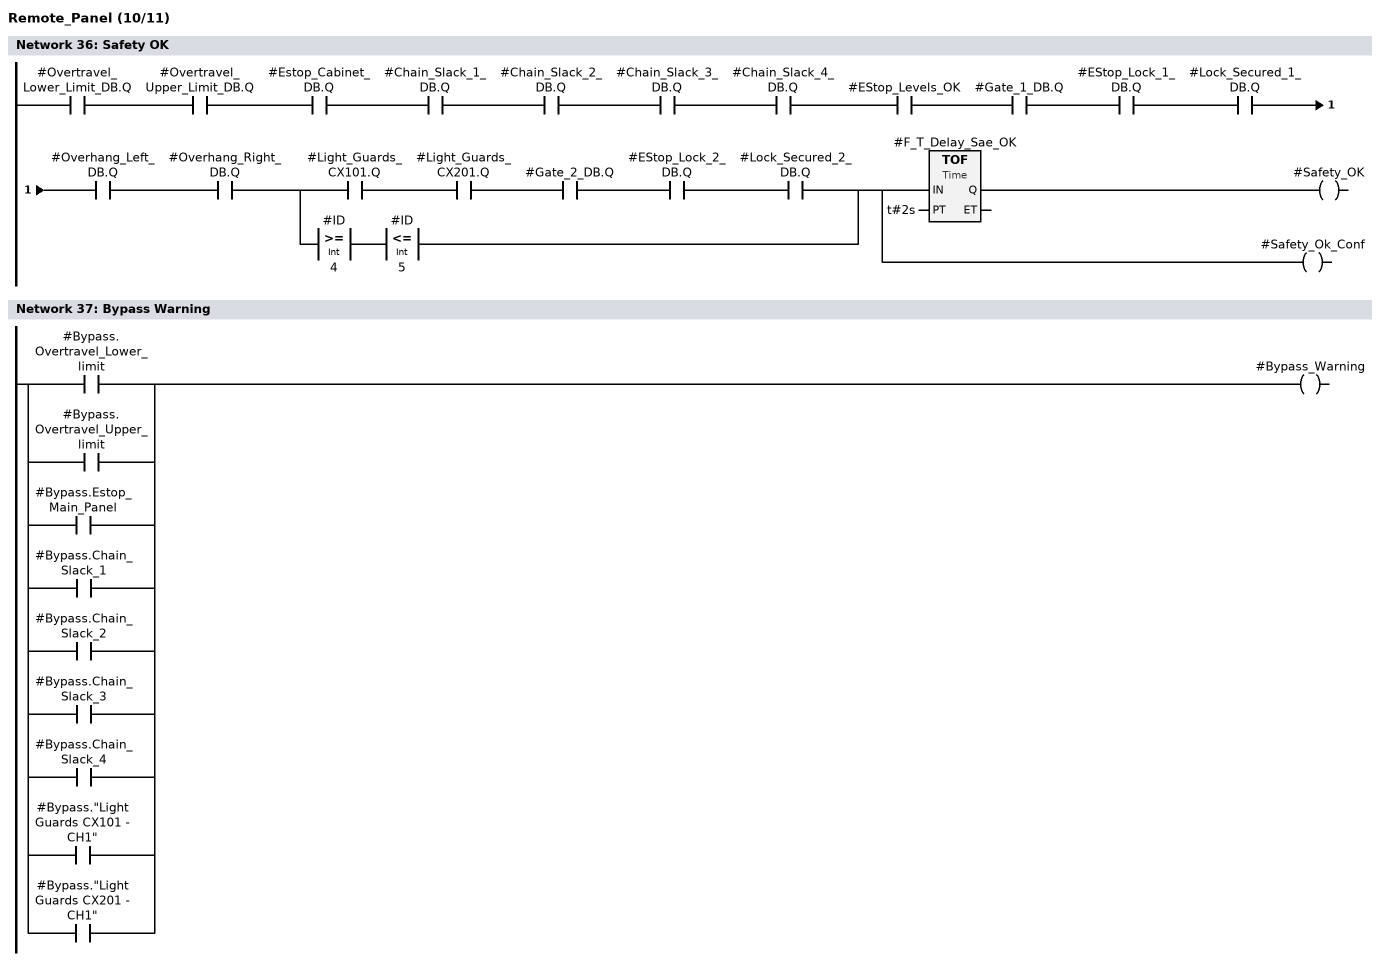
   RUNG wire#powerrail
      Contact( #Overtravel_Lower_Limit_DB.Q )
      Contact( #Overtravel_Upper_Limit_DB.Q )
      Contact( #Estop_Cabinet_DB.Q )
      Contact( #Chain_Slack_1_DB.Q )
      Contact( #Chain_Slack_2_DB.Q )
      Contact( #Chain_Slack_3_DB.Q )
      Contact( #Chain_Slack_4_DB.Q )
      Contact( #EStop_Levels_OK )
      Contact( #Gate_1_DB.Q )
      Contact( #EStop_Lock_1_DB.Q )
      Contact( #Lock_Secured_1_DB.Q )
      Contact( #Overhang_Left_DB.Q )
      Contact( #Overhang_Right_DB.Q )
      wire#w1
      Contact( #Light_Guards_CX101.Q )
      Contact( #Light_Guards_CX201.Q )
      Contact( #Gate_2_DB.Q )
      Contact( #EStop_Lock_2_DB.Q )
      Contact( #Lock_Secured_2_DB.Q )
      wire#w2
      { S7_Templates := "[time_type := Time, codedbool_type := DInt]" } #F_T_Delay_Sae_OK.TOF(pt := t#2s, et =>)
      Coil( #Safety_OK )
   END_RUNG
   RUNG wire#w1
      { S7_Templates := "SrcType := Int" } GE_Contact(in1 := #ID, in2 := 4)
      { S7_Templates := "SrcType := Int" } LE_Contact(in1 := #ID, in2 := 5)
   END_RUNG wire#w2
   RUNG wire#w2
      Coil( #Safety_Ok_Conf )
   END_RUNG
   // the same network as SCL:
   #_w1 := #Overtravel_Lower_Limit_DB.Q AND #Overtravel_Upper_Limit_DB.Q AND #Estop_Cabinet_DB.Q AND #Chain_Slack_1_DB.Q AND #Chain_Slack_2_DB.Q AND #Chain_Slack_3_DB.Q AND #Chain_Slack_4_DB.Q AND #EStop_Levels_OK AND #Gate_1_DB.Q AND #EStop_Lock_1_DB.Q AND #Lock_Secured_1_DB.Q AND #Overhang_Left_DB.Q AND #Overhang_Right_DB.Q AND ((#Light_Guards_CX101.Q AND #Light_Guards_CX201.Q AND #Gate_2_DB.Q AND #EStop_Lock_2_DB.Q AND #Lock_Secured_2_DB.Q) OR ((#ID >= 4) AND (#ID <= 5)));
   #F_T_Delay_Sae_OK.TOF(IN := #_w1, PT := t#2s);
   #Safety_OK := #F_T_Delay_Sae_OK.Q;
   #Safety_Ok_Conf := #_w1;
END_REGION

REGION Network 37: Bypass Warning
   RUNG wire#powerrail
      Contact( #Bypass.Overtravel_Lower_limit )
      wire#w1
      Coil( #Bypass_Warning )
   END_RUNG
   RUNG wire#powerrail
      Contact( #Bypass.Overtravel_Upper_limit )
   END_RUNG wire#w1
   RUNG wire#powerrail
      Contact( #Bypass.Estop_Main_Panel )
   END_RUNG wire#w1
   RUNG wire#powerrail
      Contact( #Bypass.Chain_Slack_1 )
   END_RUNG wire#w1
   RUNG wire#powerrail
      Contact( #Bypass.Chain_Slack_2 )
   END_RUNG wire#w1
   RUNG wire#powerrail
      Contact( #Bypass.Chain_Slack_3 )
   END_RUNG wire#w1
   RUNG wire#powerrail
      Contact( #Bypass.Chain_Slack_4 )
   END_RUNG wire#w1
   RUNG wire#powerrail
      Contact( #Bypass."Light Guards CX101 - CH1" )
   END_RUNG wire#w1
   RUNG wire#powerrail
      Contact( #Bypass."Light Guards CX201 - CH1" )
   END_RUNG wire#w1
   // the same network as SCL:
   #Bypass_Warning := #Bypass.Overtravel_Lower_limit OR #Bypass.Overtravel_Upper_limit OR #Bypass.Estop_Main_Panel OR #Bypass.Chain_Slack_1 OR #Bypass.Chain_Slack_2 OR #Bypass.Chain_Slack_3 OR #Bypass.Chain_Slack_4 OR #Bypass."Light Guards CX101 - CH1" OR #Bypass."Light Guards CX201 - CH1";
END_REGION

REGION Network 38: Enable outputs
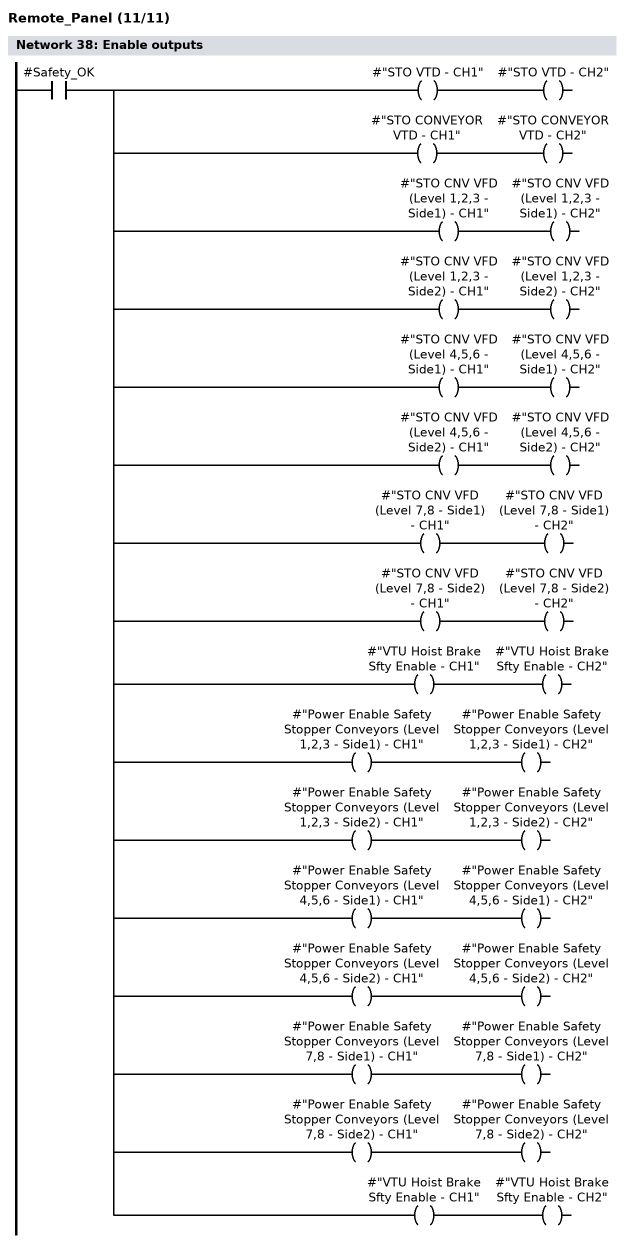
   RUNG wire#powerrail
      Contact( #Safety_OK )
      wire#w1
      Coil( #"STO VTD - CH1" )
      Coil( #"STO VTD - CH2" )
   END_RUNG
   RUNG wire#w1
      Coil( #"STO CONVEYOR VTD - CH1" )
      Coil( #"STO CONVEYOR VTD - CH2" )
   END_RUNG
   RUNG wire#w1
      Coil( #"STO CNV VFD (Level 1,2,3 - Side1) - CH1" )
      Coil( #"STO CNV VFD (Level 1,2,3 - Side1) - CH2" )
   END_RUNG
   RUNG wire#w1
      Coil( #"STO CNV VFD (Level 1,2,3 - Side2) - CH1" )
      Coil( #"STO CNV VFD (Level 1,2,3 - Side2) - CH2" )
   END_RUNG
   RUNG wire#w1
      Coil( #"STO CNV VFD (Level 4,5,6 - Side1) - CH1" )
      Coil( #"STO CNV VFD (Level 4,5,6 - Side1) - CH2" )
   END_RUNG
   RUNG wire#w1
      Coil( #"STO CNV VFD (Level 4,5,6 - Side2) - CH1" )
      Coil( #"STO CNV VFD (Level 4,5,6 - Side2) - CH2" )
   END_RUNG
   RUNG wire#w1
      Coil( #"STO CNV VFD (Level 7,8 - Side1) - CH1" )
      Coil( #"STO CNV VFD (Level 7,8 - Side1) - CH2" )
   END_RUNG
   RUNG wire#w1
      Coil( #"STO CNV VFD (Level 7,8 - Side2) - CH1" )
      Coil( #"STO CNV VFD (Level 7,8 - Side2) - CH2" )
   END_RUNG
   RUNG wire#w1
      Coil( #"VTU Hoist Brake Sfty Enable - CH1" )
      Coil( #"VTU Hoist Brake Sfty Enable - CH2" )
   END_RUNG
   RUNG wire#w1
      Coil( #"Power Enable Safety Stopper Conveyors (Level 1,2,3 - Side1) - CH1" )
      Coil( #"Power Enable Safety Stopper Conveyors (Level 1,2,3 - Side1) - CH2" )
   END_RUNG
   RUNG wire#w1
      Coil( #"Power Enable Safety Stopper Conveyors (Level 1,2,3 - Side2) - CH1" )
      Coil( #"Power Enable Safety Stopper Conveyors (Level 1,2,3 - Side2) - CH2" )
   END_RUNG
   RUNG wire#w1
      Coil( #"Power Enable Safety Stopper Conveyors (Level 4,5,6 - Side1) - CH1" )
      Coil( #"Power Enable Safety Stopper Conveyors (Level 4,5,6 - Side1) - CH2" )
   END_RUNG
   RUNG wire#w1
      Coil( #"Power Enable Safety Stopper Conveyors (Level 4,5,6 - Side2) - CH1" )
      Coil( #"Power Enable Safety Stopper Conveyors (Level 4,5,6 - Side2) - CH2" )
   END_RUNG
   RUNG wire#w1
      Coil( #"Power Enable Safety Stopper Conveyors (Level 7,8 - Side1) - CH1" )
      Coil( #"Power Enable Safety Stopper Conveyors (Level 7,8 - Side1) - CH2" )
   END_RUNG
   RUNG wire#w1
      Coil( #"Power Enable Safety Stopper Conveyors (Level 7,8 - Side2) - CH1" )
      Coil( #"Power Enable Safety Stopper Conveyors (Level 7,8 - Side2) - CH2" )
   END_RUNG
   RUNG wire#w1
      Coil( #"VTU Hoist Brake Sfty Enable - CH1" )
      Coil( #"VTU Hoist Brake Sfty Enable - CH2" )
   END_RUNG
   // the same network as SCL:
   #"STO VTD - CH1" := #Safety_OK;
   #"STO VTD - CH2" := #Safety_OK;
   #"STO CONVEYOR VTD - CH1" := #Safety_OK;
   #"STO CONVEYOR VTD - CH2" := #Safety_OK;
   #"STO CNV VFD (Level 1,2,3 - Side1) - CH1" := #Safety_OK;
   #"STO CNV VFD (Level 1,2,3 - Side1) - CH2" := #Safety_OK;
   #"STO CNV VFD (Level 1,2,3 - Side2) - CH1" := #Safety_OK;
   #"STO CNV VFD (Level 1,2,3 - Side2) - CH2" := #Safety_OK;
   #"STO CNV VFD (Level 4,5,6 - Side1) - CH1" := #Safety_OK;
   #"STO CNV VFD (Level 4,5,6 - Side1) - CH2" := #Safety_OK;
   #"STO CNV VFD (Level 4,5,6 - Side2) - CH1" := #Safety_OK;
   #"STO CNV VFD (Level 4,5,6 - Side2) - CH2" := #Safety_OK;
   #"STO CNV VFD (Level 7,8 - Side1) - CH1" := #Safety_OK;
   #"STO CNV VFD (Level 7,8 - Side1) - CH2" := #Safety_OK;
   #"STO CNV VFD (Level 7,8 - Side2) - CH1" := #Safety_OK;
   #"STO CNV VFD (Level 7,8 - Side2) - CH2" := #Safety_OK;
   #"VTU Hoist Brake Sfty Enable - CH1" := #Safety_OK;
   #"VTU Hoist Brake Sfty Enable - CH2" := #Safety_OK;
   #"Power Enable Safety Stopper Conveyors (Level 1,2,3 - Side1) - CH1" := #Safety_OK;
   #"Power Enable Safety Stopper Conveyors (Level 1,2,3 - Side1) - CH2" := #Safety_OK;
   #"Power Enable Safety Stopper Conveyors (Level 1,2,3 - Side2) - CH1" := #Safety_OK;
   #"Power Enable Safety Stopper Conveyors (Level 1,2,3 - Side2) - CH2" := #Safety_OK;
   #"Power Enable Safety Stopper Conveyors (Level 4,5,6 - Side1) - CH1" := #Safety_OK;
   #"Power Enable Safety Stopper Conveyors (Level 4,5,6 - Side1) - CH2" := #Safety_OK;
   #"Power Enable Safety Stopper Conveyors (Level 4,5,6 - Side2) - CH1" := #Safety_OK;
   #"Power Enable Safety Stopper Conveyors (Level 4,5,6 - Side2) - CH2" := #Safety_OK;
   #"Power Enable Safety Stopper Conveyors (Level 7,8 - Side1) - CH1" := #Safety_OK;
   #"Power Enable Safety Stopper Conveyors (Level 7,8 - Side1) - CH2" := #Safety_OK;
   #"Power Enable Safety Stopper Conveyors (Level 7,8 - Side2) - CH1" := #Safety_OK;
   #"Power Enable Safety Stopper Conveyors (Level 7,8 - Side2) - CH2" := #Safety_OK;
   #"VTU Hoist Brake Sfty Enable - CH1" := #Safety_OK;
   #"VTU Hoist Brake Sfty Enable - CH2" := #Safety_OK;
END_REGION
END_FUNCTION_BLOCK
